ABB RAPID module: SetProg.mod

%%%
  VERSION:1
  LANGUAGE:ENGLISH
%%%
MODULE MOD_SetProg

    ! -------------------------------
    ! Define customized variables here
    ! ...

	! Tool variables:
	PERS tooldata ToolS := [TRUE,[[10.000,20.000,150.000],[1.00000000,0.00000000,0.00000000,0.00000000]],[1,[0,0,20],[1,0,0,0],0,0,0.005]];

	! Reference variables:
	PERS wobjdata FrameS := [FALSE, TRUE, "", [[0,0,0],[1,0,0,0]],[[1234.570,-98.765,50.500],[0.96592583,0.00000000,0.00000000,0.25881905]]];

	PROC Main()
		ConfJ \On;
		ConfL \Off;
		! Program generated by RoboDK v6.0.7 for ABB IRB 120-3/0.6 on XX/XX/XXXX 12:58:42
		! Using nominal kinematics.
		MoveAbsJ [[0.000000,-10.000000,20.000000,0.000000,30.000000,0.000000],[9E+09,9E+09,9E+09,9E+09,9E+09,9E+09]],v500,z1,ToolS \WObj:=FrameS;
		MoveL [[-615.584,550.281,371.534],[0.40821789,0.23456972,0.87542610,-0.10938165],[0,0,0,0],[9E+09,9E+09,9E+09,9E+09,9E+09,9E+09]],v500,z1,ToolS \WObj:=FrameS;
		MoveC [[-618.417,609.652,333.231],[0.40821789,0.23456972,0.87542610,-0.10938165],[0,0,0,0],[9E+09,9E+09,9E+09,9E+09,9E+09,9E+09]],[[-671.251,582.420,294.929],[0.40821789,0.23456972,0.87542610,-0.10938165],[0,0,0,0],[9E+09,9E+09,9E+09,9E+09,9E+09,9E+09]],v500,z1,ToolS \WObj:=FrameS;
		MoveAbsJ [[20.000000,-10.000000,20.000000,0.000000,30.000000,0.000000],[9E+09,9E+09,9E+09,9E+09,9E+09,9E+09]],v500,z1,ToolS \WObj:=FrameS;
		WaitTime 0.250;
		MoveAbsJ [[30.000000,-20.000000,40.000000,60.000000,-45.000000,-100.000000],[9E+09,9E+09,9E+09,9E+09,9E+09,9E+09]],v500,z1,ToolS \WObj:=FrameS;
	ENDPROC

ENDMODULE
